FUNCTION_BLOCK FB_STOEBERSDS_Reset
(*

The function block used to reset an axis

Constructor: 		Patryk Panylo
Company:		E. Riexinger GmbH
Date:			22.09.2015
Version:			1.00

Date:			Revision:		Who:				Comment

*)
VAR_INPUT
	(* Input variables / Eingang Variablen *)
	bExecute					:BOOL;		(* Execut the function block *)
END_VAR
VAR_OUTPUT
	(* Output variables / Ausgang Variablen *)
	bDone						:BOOL;			(* Status = TRUE indicates that the axis is ready for operation. *)
	bBusy						:BOOL;			(* Program busy *)
	bError						:BOOL;			(* Error *)
	udnErrorNo					:UDINT;			(* Error number *)
	sErrorMsg					:STRING; 		(* Error message *)
END_VAR
VAR_IN_OUT
	(* Input Output variables / Ausgang Variablen *)
	Axis							:ST_AXIS_REF;
END_VAR
VAR
	(* Enummerations *)

	(* Variables *)

	(* References *)

	(* Interfaces *)

	(* Instances *)
	rtExecute						:R_TRIG;
END_VAR


rtExecute(CLK := bExecute);       (* Error *)

IF rtExecute.Q
THEN
	bBusy := TRUE;
	Axis.stPlcToNc.stBaseDevice.bFaultReset := TRUE;

ELSIF NOT Axis.stNcToPlc.stBaseDevice.bError      (* Error *)
THEN
	bBusy := FALSE;
	Axis.stPlcToNc.stBaseDevice.bFaultReset := FALSE;
END_IF;

bDone := bExecute
		AND NOT bBusy
		AND NOT  Axis.stNcToPlc.stBaseDevice.bError;        (* Error *)

END_FUNCTION_BLOCK

(* stored: Version 1.1.0.1, ProductVersion 3.1.4024.15
   POU FB_STOEBERSDS_Reset: Id {4e1f28c0-219b-48e3-b85f-cee91862b436}, SpecialFunc None *)
